(* PLC project Motor_StartStop_TM241CE24T, PLCAutoPilot M241 Generator 2.0 *)
(* stored: creationDateTime 2025-12-30T00:00:00, modificationDateTime 2025-12-30T00:00:00 *)

PROGRAM GVL
  VAR_GLOBAL
    StartPB AT %IX0.0 : BOOL;  (* Start Pushbutton (NO) *)
    StopPB AT %IX0.1 : BOOL;  (* Stop Pushbutton (NC) *)
    OverloadTrip AT %IX0.2 : BOOL;  (* Thermal Overload Relay (NC) *)
    EmergencyStop AT %IX0.3 : BOOL;  (* Emergency Stop (NC) *)
    MotorContactor AT %QX0.0 : BOOL;  (* Main Contactor K1 *)
    RunIndicator AT %QX0.1 : BOOL;  (* Run Indicator Lamp *)
    FaultIndicator AT %QX0.2 : BOOL;  (* Fault Indicator Lamp *)
  END_VAR

END_PROGRAM

(* Motor Start/Stop Control for TM241CE24T INPUTS: - StartPB (%IX0.0): Start pushbutton (NO) - StopPB (%IX0.1): Stop pushbutton (NC) - OverloadTrip (%IX0.2): Thermal overload relay (NC) - EmergencyStop (%IX0.3): Emergency stop (NC) OUTPUTS: - MotorContactor (%QX0.0): Main contactor K1 - RunIndicator (%QX0.1): Run indicator lamp - FaultIndicator (%QX0.2): Fault indicator lamp FEATURES: - 3 second startup delay (anti-chatter) - Overload fault latching with reset - Emergency stop interlock - Run and fault indication Generated by PLCAutoPilot *)
PROGRAM Motor_Control
  VAR
    MotorRunning : BOOL;  (* Motor Running Status *)
    MotorFault : BOOL;  (* Motor Fault Latched *)
    StartupTimer : TON;  (* 3 second startup delay *)
    SafetyOK : BOOL;  (* All safety conditions met *)
  END_VAR
  VAR  (* added by the conversion: wires and edge detectors of the diagram *)
    _AND1_OUT : BOOL;
    _AND20_OUT : BOOL;
    _TON30_ET : ANY;
    _TON30_OUT : BOOL;
    _OR50_OUT : BOOL;
    _SR40_OUT : BOOL;
    _RS70_OUT : BOOL;
  END_VAR

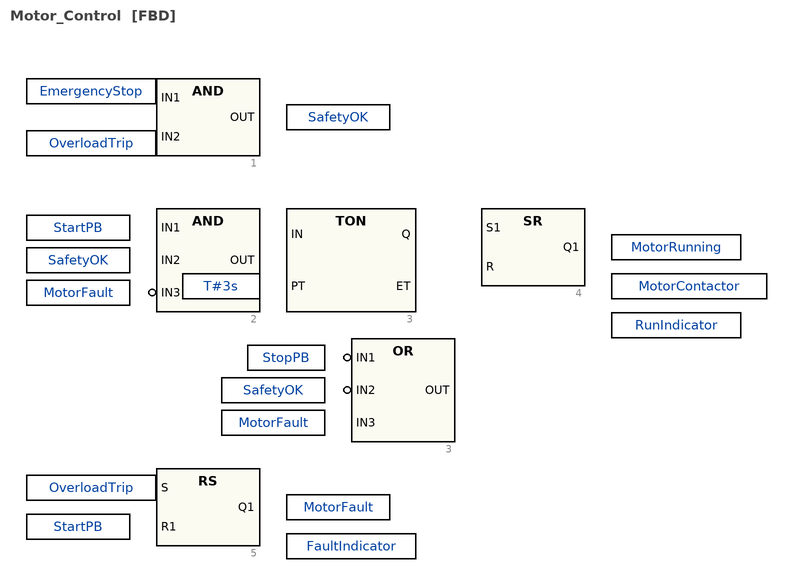
(* FBD diagram, written out as Structured Text *)
_AND1_OUT := EmergencyStop AND NOT OverloadTrip;
_AND20_OUT := StartPB AND SafetyOK AND NOT MotorFault;
_TON30_OUT := TON(IN := _AND20_OUT, PT := T#3s, ET => _TON30_ET);
_OR50_OUT := NOT StopPB OR NOT SafetyOK OR MotorFault;
_SR40_OUT := SR(_TON30_OUT, _OR50_OUT);
_RS70_OUT := RS(OverloadTrip, StartPB);
SafetyOK := _AND1_OUT;
MotorRunning := _SR40_OUT;
MotorContactor := _SR40_OUT;
RunIndicator := _SR40_OUT;
MotorFault := _RS70_OUT;
FaultIndicator := _RS70_OUT;
END_PROGRAM

CONFIGURATION TM241CE24T
  RESOURCE Application ON PLC
    TASK MAST(INTERVAL := T#20ms, PRIORITY := 1);
    PROGRAM Motor_Control_Instance WITH MAST : Motor_Control;
  END_RESOURCE
END_CONFIGURATION
